Staubli VAL3: getlog.pgx

public program getlog(string& x_sLog[], num x_nType)
  local num i
  local num j
begin
  for i=0 to size(x_sLog)-1
    //获取当前日志
    //如果是类型0，表示筛选全部类型的日志，如果是其他类型，则根据当前的日志类型筛选
    if x_nType==0
      x_sLog[i]=sLog[sel(nIndex-1-i>=0,nIndex-1-i,nIndex-1-i+size(sLog))]
    else
      //筛选需要的类型
      while nLogType[sel(nIndex-1-j>=0,nIndex-1-j,nIndex-1-j+size(sLog))]!=x_nType and j<size(sLog)
        j=j+1
      endWhile
      //超过了全部日志数组的大小，说明遍历了一遍，则跳出
      if j>=size(sLog)
        return
      endIf
      x_sLog[i]=sLog[sel(nIndex-1-j>=0,nIndex-1-j,nIndex-1-j+size(sLog))]
      j=j+1
    endIf
  endFor
end
